Fanuc KAREL source: kb00048.KL

PROGRAM KB00048
%NOLOCKGROUP
VAR
P1:REAL;RESULT:REAL
BEGIN
--
P1=1.0
RESULT=COS(P1)
END KB00048
